(*
SPDX-FileCopyrightText: © 2026 Oleksandr Tiutyk <trofimich@gmail.com>
SPDX-License-Identifier: MIT
License: https://opensource.org/license/mit
*)

{attribute 'qualified_only'}
VAR_GLOBAL
	Name : STRING := 'TOF_Tests';
END_VAR

(* stored: Version 1.1.0.1
   GVL CurrentNamespace: Id {a2446931-0eaa-4b6b-b048-aef391c46fe6} *)
